// TIA Portal V19 export
DATA_BLOCK "V20_BLOCK_DB"   // DB83
// stored: InstanceOfName V20_BLOCK, InstanceOfType FB
"V20_BLOCK"
   // VAR
   //    MB_LOAD { S7_SetPoint := 'True'} : Modbus_Comm_Load;
   //    MB_READ_ZSW { S7_SetPoint := 'True'} : Modbus_Master;
   //    MB_READ_HIW { S7_SetPoint := 'True'} : Modbus_Master;
   //    MB_WRITE_STW { S7_SetPoint := 'True'} : Modbus_Master;
   //    MB_WRITE_HSW { S7_SetPoint := 'True'} : Modbus_Master;
   //    DRIVE { S7_SetPoint := 'True'} : Array[1..11] of "VFD";
   //    DRIVE_ID { S7_SetPoint := 'True'} : Int;
   //    STATUS : Int;
   //    MB_DB : P2P_MB_BASE;
   //    ZSW_DELAY { S7_SetPoint := 'True'} : TON_TIME;
   //    HIW_DELAY { S7_SetPoint := 'True'} : TON_TIME;
   //    STW_DELAY { S7_SetPoint := 'True'} : TON_TIME;
   //    HSW_DELAY { S7_SetPoint := 'True'} : TON_TIME;
   //    MB_READ_DI { S7_SetPoint := 'True'} : Modbus_Master;
   //    Modbus_Master_Instance { S7_SetPoint := 'True'} : Modbus_Master;
   // END_VAR
BEGIN
   DRIVE[7].ADDR := 7;
   DRIVE[8].ADDR := 8;
   DRIVE[9].ADDR := 9;
   DRIVE[10].ADDR := 10;
   DRIVE[11].ADDR := 11;
END_DATA_BLOCK
